RoboDK station: Car_Painting_Model .rdk

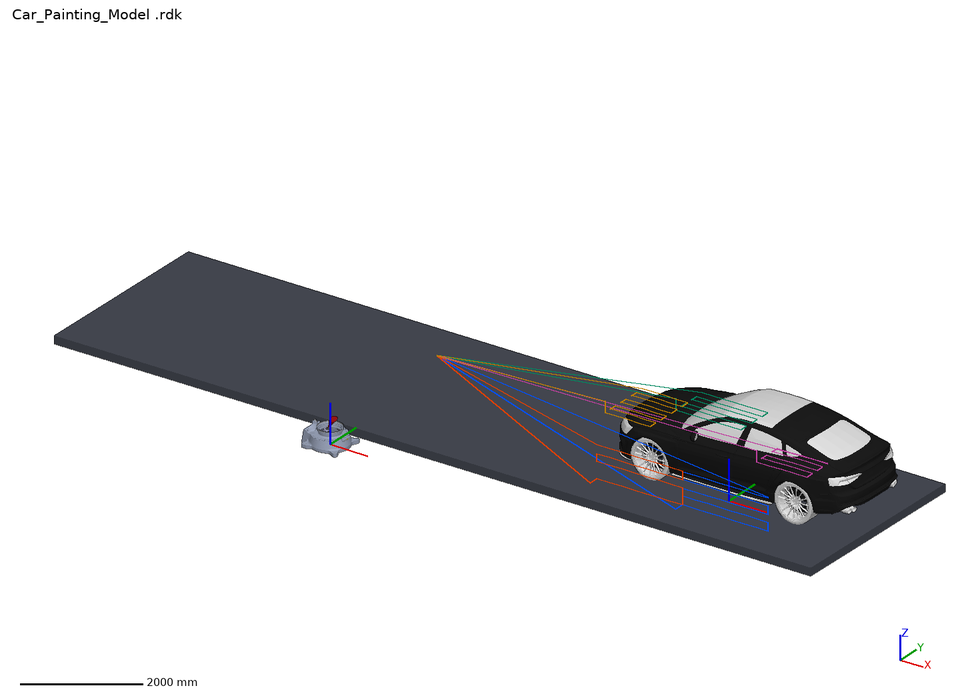
[picture v0: the station drawn from its stored meshes, robots at their saved joint values, targets as dots, program paths as lines]
Station Car_Painting_Model  (saved by RoboDK 6.0.6). Poses are relative to the parent item; angles as X-Y-Z fixed-axis rotations.
Station parameters (name, value as stored): LIN64
  - frame Comau Smart5 NJ 130-2.6 Base at (-637.82, 0, 0) mm
    - robot Comau Smart5 NJ 130-2.6: 6 axes, payload 130 kg, reach 2616 mm, repeatability 0.07 mm, weight 1050 kg
        joint limits [-180, -75, -351, -280, -120, -720] to [180, 95, 170, 280, 120, 720]; home [0, 0, -90, 0, 0, 0]; saved at [0, 0, -90, 0, 0, 0]
      - tool Generic Paint Sprayer, TCP at (50, 0, 450) mm, rotated rx 0 ry 30 rz 0 deg, size 277.6 x 203.2 x 501.7 mm
  - frame CarFrame at (5862.18, 2000, 0) mm
    - object CAN_CAR_BLEND_V12 at (230.98, 0, 65.42) mm, rotated rx 80 ry 0 rz 90 deg, size 2096.9 x 1491.7 x 4800 mm, geometry from CAN_CAR_BLEND_V12.glb
    - target CHK_Nose (Cartesian target) at (2400, 0, 600) mm; joints [0, 0, -90, 0, 0, 0] of Comau Smart5 NJ 130-2.6
    - target CHK_Tail (Cartesian target) at (-2400, 0, 600) mm; joints [0, 0, -90, 0, 0, 0] of Comau Smart5 NJ 130-2.6
    - target CHK_Left_door (Cartesian target) at (0, 1048.43, 800) mm; joints [0, 0, -90, 0, 0, 0] of Comau Smart5 NJ 130-2.6
    - target CHK_Right_door (Cartesian target) at (0, -1048.43, 800) mm; joints [0, 0, -90, 0, 0, 0] of Comau Smart5 NJ 130-2.6
    - target CHK_Roof (Cartesian target) at (0, 0, 1491.68) mm; joints [0, 0, -90, 0, 0, 0] of Comau Smart5 NJ 130-2.6
    - target P_Home (joint target) at (-4384.42, -2000, 2190) mm, rotated rx 180 ry 60 rz 180 deg; joints [0, 0, -90, 0, 0, 0] of Comau Smart5 NJ 130-2.6
    - target P_Right_Front_J_approach (Cartesian target) at (0, -1498.5, 450) mm, rotated rx -90 ry 0 rz 0 deg; joints [0, 0, -90, 0, 0, 0] of Comau Smart5 NJ 130-2.6
    - target P_Right_Front_J_p00_w00 (Cartesian target) at (0, -1298.5, 450) mm, rotated rx -90 ry 0 rz 0 deg; joints [0, 0, -90, 0, 0, 0] of Comau Smart5 NJ 130-2.6
    - target P_Right_Front_J_p00_w01 (Cartesian target) at (242.86, -1298.5, 450) mm, rotated rx -90 ry 0 rz 0 deg; joints [0, 0, -90, 0, 0, 0] of Comau Smart5 NJ 130-2.6
    - target P_Right_Front_J_p00_w02 (Cartesian target) at (485.71, -1298.5, 450) mm, rotated rx -90 ry 0 rz 0 deg; joints [0, 0, -90, 0, 0, 0] of Comau Smart5 NJ 130-2.6
    - target P_Right_Front_J_p00_w03 (Cartesian target) at (728.57, -1298.5, 450) mm, rotated rx -90 ry 0 rz 0 deg; joints [0, 0, -90, 0, 0, 0] of Comau Smart5 NJ 130-2.6
    - target P_Right_Front_J_p00_w04 (Cartesian target) at (971.43, -1298.5, 450) mm, rotated rx -90 ry 0 rz 0 deg; joints [0, 0, -90, 0, 0, 0] of Comau Smart5 NJ 130-2.6
    - target P_Right_Front_J_p00_w05 (Cartesian target) at (1214.29, -1298.5, 450) mm, rotated rx -90 ry 0 rz 0 deg; joints [0, 0, -90, 0, 0, 0] of Comau Smart5 NJ 130-2.6
    - target P_Right_Front_J_p00_w06 (Cartesian target) at (1457.14, -1298.5, 450) mm, rotated rx -90 ry 0 rz 0 deg; joints [0, 0, -90, 0, 0, 0] of Comau Smart5 NJ 130-2.6
    - target P_Right_Front_J_p00_w07 (Cartesian target) at (1700, -1298.5, 450) mm, rotated rx -90 ry 0 rz 0 deg; joints [0, 0, -90, 0, 0, 0] of Comau Smart5 NJ 130-2.6
    - target P_Right_Front_J_p01_w00 (Cartesian target) at (1700, -1298.5, 600) mm, rotated rx 90 ry 0 rz 180 deg; joints [0, 0, -90, 0, 0, 0] of Comau Smart5 NJ 130-2.6
    - target P_Right_Front_J_p01_w01 (Cartesian target) at (1457.14, -1298.5, 600) mm, rotated rx 90 ry 0 rz 180 deg; joints [0, 0, -90, 0, 0, 0] of Comau Smart5 NJ 130-2.6
    - target P_Right_Front_J_p01_w02 (Cartesian target) at (1214.29, -1298.5, 600) mm, rotated rx 90 ry 0 rz 180 deg; joints [0, 0, -90, 0, 0, 0] of Comau Smart5 NJ 130-2.6
    - target P_Right_Front_J_p01_w03 (Cartesian target) at (971.43, -1298.5, 600) mm, rotated rx 90 ry 0 rz 180 deg; joints [0, 0, -90, 0, 0, 0] of Comau Smart5 NJ 130-2.6
    - target P_Right_Front_J_p01_w04 (Cartesian target) at (728.57, -1298.5, 600) mm, rotated rx 90 ry 0 rz 180 deg; joints [0, 0, -90, 0, 0, 0] of Comau Smart5 NJ 130-2.6
    - target P_Right_Front_J_p01_w05 (Cartesian target) at (485.71, -1298.5, 600) mm, rotated rx 90 ry 0 rz 180 deg; joints [0, 0, -90, 0, 0, 0] of Comau Smart5 NJ 130-2.6
    - target P_Right_Front_J_p01_w06 (Cartesian target) at (242.86, -1298.5, 600) mm, rotated rx 90 ry 0 rz 180 deg; joints [0, 0, -90, 0, 0, 0] of Comau Smart5 NJ 130-2.6
    - target P_Right_Front_J_p01_w07 (Cartesian target) at (0, -1298.5, 600) mm, rotated rx 90 ry 0 rz 180 deg; joints [0, 0, -90, 0, 0, 0] of Comau Smart5 NJ 130-2.6
    - target P_Right_Front_J_p02_w00 (Cartesian target) at (0, -1298.5, 750) mm, rotated rx -90 ry 0 rz 0 deg; joints [0, 0, -90, 0, 0, 0] of Comau Smart5 NJ 130-2.6
    - target P_Right_Front_J_p02_w01 (Cartesian target) at (242.86, -1298.5, 750) mm, rotated rx -90 ry 0 rz 0 deg; joints [0, 0, -90, 0, 0, 0] of Comau Smart5 NJ 130-2.6
    - target P_Right_Front_J_p02_w02 (Cartesian target) at (485.71, -1298.5, 750) mm, rotated rx -90 ry 0 rz 0 deg; joints [0, 0, -90, 0, 0, 0] of Comau Smart5 NJ 130-2.6
    - target P_Right_Front_J_p02_w03 (Cartesian target) at (728.57, -1298.5, 750) mm, rotated rx -90 ry 0 rz 0 deg; joints [0, 0, -90, 0, 0, 0] of Comau Smart5 NJ 130-2.6
    - target P_Right_Front_J_p02_w04 (Cartesian target) at (971.43, -1298.5, 750) mm, rotated rx -90 ry 0 rz 0 deg; joints [0, 0, -90, 0, 0, 0] of Comau Smart5 NJ 130-2.6
    - target P_Right_Front_J_p02_w05 (Cartesian target) at (1214.29, -1298.5, 750) mm, rotated rx -90 ry 0 rz 0 deg; joints [0, 0, -90, 0, 0, 0] of Comau Smart5 NJ 130-2.6
    - target P_Right_Front_J_p02_w06 (Cartesian target) at (1457.14, -1298.5, 750) mm, rotated rx -90 ry 0 rz 0 deg; joints [0, 0, -90, 0, 0, 0] of Comau Smart5 NJ 130-2.6
    - target P_Right_Front_J_p02_w07 (Cartesian target) at (1700, -1298.5, 750) mm, rotated rx -90 ry 0 rz 0 deg; joints [0, 0, -90, 0, 0, 0] of Comau Smart5 NJ 130-2.6
    - target P_Right_Front_J_p03_w00 (Cartesian target) at (1700, -1298.5, 900) mm, rotated rx 90 ry 0 rz 180 deg; joints [0, 0, -90, 0, 0, 0] of Comau Smart5 NJ 130-2.6
    - target P_Right_Front_J_p03_w01 (Cartesian target) at (1457.14, -1298.5, 900) mm, rotated rx 90 ry 0 rz 180 deg; joints [0, 0, -90, 0, 0, 0] of Comau Smart5 NJ 130-2.6
    - target P_Right_Front_J_p03_w02 (Cartesian target) at (1214.29, -1298.5, 900) mm, rotated rx 90 ry 0 rz 180 deg; joints [0, 0, -90, 0, 0, 0] of Comau Smart5 NJ 130-2.6
    - target P_Right_Front_J_p03_w03 (Cartesian target) at (971.43, -1298.5, 900) mm, rotated rx 90 ry 0 rz 180 deg; joints [0, 0, -90, 0, 0, 0] of Comau Smart5 NJ 130-2.6
    - target P_Right_Front_J_p03_w04 (Cartesian target) at (728.57, -1298.5, 900) mm, rotated rx 90 ry 0 rz 180 deg; joints [0, 0, -90, 0, 0, 0] of Comau Smart5 NJ 130-2.6
    - target P_Right_Front_J_p03_w05 (Cartesian target) at (485.71, -1298.5, 900) mm, rotated rx 90 ry 0 rz 180 deg; joints [0, 0, -90, 0, 0, 0] of Comau Smart5 NJ 130-2.6
    - target P_Right_Front_J_p03_w06 (Cartesian target) at (242.86, -1298.5, 900) mm, rotated rx 90 ry 0 rz 180 deg; joints [0, 0, -90, 0, 0, 0] of Comau Smart5 NJ 130-2.6
    - target P_Right_Front_J_p03_w07 (Cartesian target) at (0, -1298.5, 900) mm, rotated rx 90 ry 0 rz 180 deg; joints [0, 0, -90, 0, 0, 0] of Comau Smart5 NJ 130-2.6
    - target P_Right_Front_J_p04_w00 (Cartesian target) at (0, -1298.5, 1050) mm, rotated rx -90 ry 0 rz 0 deg; joints [0, 0, -90, 0, 0, 0] of Comau Smart5 NJ 130-2.6
    - target P_Right_Front_J_p04_w01 (Cartesian target) at (242.86, -1298.5, 1050) mm, rotated rx -90 ry 0 rz 0 deg; joints [0, 0, -90, 0, 0, 0] of Comau Smart5 NJ 130-2.6
    - target P_Right_Front_J_p04_w02 (Cartesian target) at (485.71, -1298.5, 1050) mm, rotated rx -90 ry 0 rz 0 deg; joints [0, 0, -90, 0, 0, 0] of Comau Smart5 NJ 130-2.6
    - target P_Right_Front_J_p04_w03 (Cartesian target) at (728.57, -1298.5, 1050) mm, rotated rx -90 ry 0 rz 0 deg; joints [0, 0, -90, 0, 0, 0] of Comau Smart5 NJ 130-2.6
    - target P_Right_Front_J_p04_w04 (Cartesian target) at (971.43, -1298.5, 1050) mm, rotated rx -90 ry 0 rz 0 deg; joints [0, 0, -90, 0, 0, 0] of Comau Smart5 NJ 130-2.6
    - target P_Right_Front_J_p04_w05 (Cartesian target) at (1214.29, -1298.5, 1050) mm, rotated rx -90 ry 0 rz 0 deg; joints [0, 0, -90, 0, 0, 0] of Comau Smart5 NJ 130-2.6
    - target P_Right_Front_J_p04_w06 (Cartesian target) at (1457.14, -1298.5, 1050) mm, rotated rx -90 ry 0 rz 0 deg; joints [0, 0, -90, 0, 0, 0] of Comau Smart5 NJ 130-2.6
    - target P_Right_Front_J_p04_w07 (Cartesian target) at (1700, -1298.5, 1050) mm, rotated rx -90 ry 0 rz 0 deg; joints [0, 0, -90, 0, 0, 0] of Comau Smart5 NJ 130-2.6
    - target P_Right_Rear_J_approach (Cartesian target) at (-1700, -1498.5, 450) mm, rotated rx -90 ry 0 rz 0 deg; joints [-106.937, 43.545, -212.911, 92.647, 99.906, 63.406] of Comau Smart5 NJ 130-2.6
    - target P_Right_Rear_J_p00_w00 (Cartesian target) at (-1700, -1298.5, 450) mm, rotated rx -90 ry 0 rz 0 deg; joints [-106.937, 43.545, -212.911, 92.647, 99.906, 63.406] of Comau Smart5 NJ 130-2.6
    - target P_Right_Rear_J_p00_w01 (Cartesian target) at (-1457.14, -1298.5, 450) mm, rotated rx -90 ry 0 rz 0 deg; joints [-106.937, 43.545, -212.911, 92.647, 99.906, 63.406] of Comau Smart5 NJ 130-2.6
    - target P_Right_Rear_J_p00_w02 (Cartesian target) at (-1214.29, -1298.5, 450) mm, rotated rx -90 ry 0 rz 0 deg; joints [-106.937, 43.545, -212.911, 92.647, 99.906, 63.406] of Comau Smart5 NJ 130-2.6
    - target P_Right_Rear_J_p00_w03 (Cartesian target) at (-971.43, -1298.5, 450) mm, rotated rx -90 ry 0 rz 0 deg; joints [-106.937, 43.545, -212.911, 92.647, 99.906, 63.406] of Comau Smart5 NJ 130-2.6
    - target P_Right_Rear_J_p00_w04 (Cartesian target) at (-728.57, -1298.5, 450) mm, rotated rx -90 ry 0 rz 0 deg; joints [-106.937, 43.545, -212.911, 92.647, 99.906, 63.406] of Comau Smart5 NJ 130-2.6
    - target P_Right_Rear_J_p00_w05 (Cartesian target) at (-485.71, -1298.5, 450) mm, rotated rx -90 ry 0 rz 0 deg; joints [-106.937, 43.545, -212.911, 92.647, 99.906, 63.406] of Comau Smart5 NJ 130-2.6
    - target P_Right_Rear_J_p00_w06 (Cartesian target) at (-242.86, -1298.5, 450) mm, rotated rx -90 ry 0 rz 0 deg; joints [-106.937, 43.545, -212.911, 92.647, 99.906, 63.406] of Comau Smart5 NJ 130-2.6
    - target P_Right_Rear_J_p00_w07 (Cartesian target) at (0, -1298.5, 450) mm, rotated rx -90 ry 0 rz 0 deg; joints [-106.937, 43.545, -212.911, 92.647, 99.906, 63.406] of Comau Smart5 NJ 130-2.6
    - target P_Right_Rear_J_p01_w00 (Cartesian target) at (0, -1298.5, 750) mm, rotated rx -90 ry 0 rz 0 deg; joints [-106.937, 43.545, -212.911, 92.647, 99.906, 63.406] of Comau Smart5 NJ 130-2.6
    - target P_Right_Rear_J_p01_w01 (Cartesian target) at (-242.86, -1298.5, 750) mm, rotated rx -90 ry 0 rz 0 deg; joints [-106.937, 43.545, -212.911, 92.647, 99.906, 63.406] of Comau Smart5 NJ 130-2.6
    - target P_Right_Rear_J_p01_w02 (Cartesian target) at (-485.71, -1298.5, 750) mm, rotated rx -90 ry 0 rz 0 deg; joints [-106.937, 43.545, -212.911, 92.647, 99.906, 63.406] of Comau Smart5 NJ 130-2.6
    - target P_Right_Rear_J_p01_w03 (Cartesian target) at (-728.57, -1298.5, 750) mm, rotated rx -90 ry 0 rz 0 deg; joints [-106.937, 43.545, -212.911, 92.647, 99.906, 63.406] of Comau Smart5 NJ 130-2.6
    - target P_Right_Rear_J_p01_w04 (Cartesian target) at (-971.43, -1298.5, 750) mm, rotated rx -90 ry 0 rz 0 deg; joints [-106.937, 43.545, -212.911, 92.647, 99.906, 63.406] of Comau Smart5 NJ 130-2.6
    - target P_Right_Rear_J_p01_w05 (Cartesian target) at (-1214.29, -1298.5, 750) mm, rotated rx -90 ry 0 rz 0 deg; joints [-106.937, 43.545, -212.911, 92.647, 99.906, 63.406] of Comau Smart5 NJ 130-2.6
    - target P_Right_Rear_J_p01_w06 (Cartesian target) at (-1457.14, -1298.5, 750) mm, rotated rx -90 ry 0 rz 0 deg; joints [-106.937, 43.545, -212.911, 92.647, 99.906, 63.406] of Comau Smart5 NJ 130-2.6
    - target P_Right_Rear_J_p01_w07 (Cartesian target) at (-1700, -1298.5, 750) mm, rotated rx -90 ry 0 rz 0 deg; joints [-106.937, 43.545, -212.911, 92.647, 99.906, 63.406] of Comau Smart5 NJ 130-2.6
    - target P_Right_Rear_J_p02_w00 (Cartesian target) at (-1700, -1298.5, 900) mm, rotated rx 90 ry 0 rz 180 deg; joints [-106.937, 43.545, -212.911, 92.647, 99.906, 63.406] of Comau Smart5 NJ 130-2.6
    - target P_Right_Rear_J_p02_w01 (Cartesian target) at (-1457.14, -1298.5, 900) mm, rotated rx 90 ry 0 rz 180 deg; joints [-106.937, 43.545, -212.911, 92.647, 99.906, 63.406] of Comau Smart5 NJ 130-2.6
    - target P_Right_Rear_J_p02_w02 (Cartesian target) at (-1214.29, -1298.5, 900) mm, rotated rx 90 ry 0 rz 180 deg; joints [-106.937, 43.545, -212.911, 92.647, 99.906, 63.406] of Comau Smart5 NJ 130-2.6
    - target P_Right_Rear_J_p02_w03 (Cartesian target) at (-971.43, -1298.5, 900) mm, rotated rx 90 ry 0 rz 180 deg; joints [-106.937, 43.545, -212.911, 92.647, 99.906, 63.406] of Comau Smart5 NJ 130-2.6
    - target P_Right_Rear_J_p02_w04 (Cartesian target) at (-728.57, -1298.5, 900) mm, rotated rx 90 ry 0 rz 180 deg; joints [-106.937, 43.545, -212.911, 92.647, 99.906, 63.406] of Comau Smart5 NJ 130-2.6
    - target P_Right_Rear_J_p02_w05 (Cartesian target) at (-485.71, -1298.5, 900) mm, rotated rx 90 ry 0 rz 180 deg; joints [-106.937, 43.545, -212.911, 92.647, 99.906, 63.406] of Comau Smart5 NJ 130-2.6
    - target P_Right_Rear_J_p02_w06 (Cartesian target) at (-242.86, -1298.5, 900) mm, rotated rx 90 ry 0 rz 180 deg; joints [-106.937, 43.545, -212.911, 92.647, 99.906, 63.406] of Comau Smart5 NJ 130-2.6
    - target P_Right_Rear_J_p02_w07 (Cartesian target) at (0, -1298.5, 900) mm, rotated rx 90 ry 0 rz 180 deg; joints [-106.937, 43.545, -212.911, 92.647, 99.906, 63.406] of Comau Smart5 NJ 130-2.6
    - target P_Right_Rear_J_p03_w00 (Cartesian target) at (0, -1298.5, 1050) mm, rotated rx -90 ry 0 rz 0 deg; joints [-106.937, 43.545, -212.911, 92.647, 99.906, 63.406] of Comau Smart5 NJ 130-2.6
    - target P_Right_Rear_J_p03_w01 (Cartesian target) at (-242.86, -1298.5, 1050) mm, rotated rx -90 ry 0 rz 0 deg; joints [-106.937, 43.545, -212.911, 92.647, 99.906, 63.406] of Comau Smart5 NJ 130-2.6
    - target P_Right_Rear_J_p03_w02 (Cartesian target) at (-485.71, -1298.5, 1050) mm, rotated rx -90 ry 0 rz 0 deg; joints [-106.937, 43.545, -212.911, 92.647, 99.906, 63.406] of Comau Smart5 NJ 130-2.6
    - target P_Right_Rear_J_p03_w03 (Cartesian target) at (-728.57, -1298.5, 1050) mm, rotated rx -90 ry 0 rz 0 deg; joints [-106.937, 43.545, -212.911, 92.647, 99.906, 63.406] of Comau Smart5 NJ 130-2.6
    - target P_Right_Rear_J_p03_w04 (Cartesian target) at (-971.43, -1298.5, 1050) mm, rotated rx -90 ry 0 rz 0 deg; joints [-106.937, 43.545, -212.911, 92.647, 99.906, 63.406] of Comau Smart5 NJ 130-2.6
    - target P_Right_Rear_J_p03_w05 (Cartesian target) at (-1214.29, -1298.5, 1050) mm, rotated rx -90 ry 0 rz 0 deg; joints [-106.937, 43.545, -212.911, 92.647, 99.906, 63.406] of Comau Smart5 NJ 130-2.6
    - target P_Right_Rear_J_p03_w06 (Cartesian target) at (-1457.14, -1298.5, 1050) mm, rotated rx -90 ry 0 rz 0 deg; joints [-106.937, 43.545, -212.911, 92.647, 99.906, 63.406] of Comau Smart5 NJ 130-2.6
    - target P_Right_Rear_J_p03_w07 (Cartesian target) at (-1700, -1298.5, 1050) mm, rotated rx -90 ry 0 rz 0 deg; joints [-106.937, 43.545, -212.911, 92.647, 99.906, 63.406] of Comau Smart5 NJ 130-2.6
    - target P_Roof_J_approach (Cartesian target) at (-600, -648.5, 1942) mm, rotated rx 180 ry 0 rz 0 deg; joints [0, 0, -90, 0, 0, 0] of Comau Smart5 NJ 130-2.6
    - target P_Roof_J_p00_w00 (Cartesian target) at (-600, -648.5, 1742) mm, rotated rx 180 ry 0 rz 0 deg; joints [0, 0, -90, 0, 0, 0] of Comau Smart5 NJ 130-2.6
    - target P_Roof_J_p00_w01 (Cartesian target) at (-383.33, -648.5, 1742) mm, rotated rx 180 ry 0 rz 0 deg; joints [0, 0, -90, 0, 0, 0] of Comau Smart5 NJ 130-2.6
    - target P_Roof_J_p00_w02 (Cartesian target) at (-166.67, -648.5, 1742) mm, rotated rx 180 ry 0 rz 0 deg; joints [0, 0, -90, 0, 0, 0] of Comau Smart5 NJ 130-2.6
    - target P_Roof_J_p00_w03 (Cartesian target) at (50, -648.5, 1742) mm, rotated rx 180 ry 0 rz 0 deg; joints [0, 0, -90, 0, 0, 0] of Comau Smart5 NJ 130-2.6
    - target P_Roof_J_p00_w04 (Cartesian target) at (266.67, -648.5, 1742) mm, rotated rx 180 ry 0 rz 0 deg; joints [0, 0, -90, 0, 0, 0] of Comau Smart5 NJ 130-2.6
    - target P_Roof_J_p00_w05 (Cartesian target) at (483.33, -648.5, 1742) mm, rotated rx 180 ry 0 rz 0 deg; joints [0, 0, -90, 0, 0, 0] of Comau Smart5 NJ 130-2.6
    - target P_Roof_J_p00_w06 (Cartesian target) at (700, -648.5, 1742) mm, rotated rx 180 ry 0 rz 0 deg; joints [0, 0, -90, 0, 0, 0] of Comau Smart5 NJ 130-2.6
    - target P_Roof_J_p01_w00 (Cartesian target) at (700, -498.5, 1742) mm, rotated rx 180 ry 0 rz 180 deg; joints [0, 0, -90, 0, 0, 0] of Comau Smart5 NJ 130-2.6
    - target P_Roof_J_p01_w01 (Cartesian target) at (483.33, -498.5, 1742) mm, rotated rx 180 ry 0 rz 180 deg; joints [0, 0, -90, 0, 0, 0] of Comau Smart5 NJ 130-2.6
    - target P_Roof_J_p01_w02 (Cartesian target) at (266.67, -498.5, 1742) mm, rotated rx 180 ry 0 rz 180 deg; joints [0, 0, -90, 0, 0, 0] of Comau Smart5 NJ 130-2.6
    - target P_Roof_J_p01_w03 (Cartesian target) at (50, -498.5, 1742) mm, rotated rx 180 ry 0 rz 180 deg; joints [0, 0, -90, 0, 0, 0] of Comau Smart5 NJ 130-2.6
    - target P_Roof_J_p01_w04 (Cartesian target) at (-166.67, -498.5, 1742) mm, rotated rx 180 ry 0 rz 180 deg; joints [0, 0, -90, 0, 0, 0] of Comau Smart5 NJ 130-2.6
    - target P_Roof_J_p01_w05 (Cartesian target) at (-383.33, -498.5, 1742) mm, rotated rx 180 ry 0 rz 180 deg; joints [0, 0, -90, 0, 0, 0] of Comau Smart5 NJ 130-2.6
    - target P_Roof_J_p01_w06 (Cartesian target) at (-600, -498.5, 1742) mm, rotated rx 180 ry 0 rz 180 deg; joints [0, 0, -90, 0, 0, 0] of Comau Smart5 NJ 130-2.6
    - target P_Roof_J_p02_w00 (Cartesian target) at (-600, -348.5, 1742) mm, rotated rx 180 ry 0 rz 0 deg; joints [0, 0, -90, 0, 0, 0] of Comau Smart5 NJ 130-2.6
    - target P_Roof_J_p02_w01 (Cartesian target) at (-383.33, -348.5, 1742) mm, rotated rx 180 ry 0 rz 0 deg; joints [0, 0, -90, 0, 0, 0] of Comau Smart5 NJ 130-2.6
    - target P_Roof_J_p02_w02 (Cartesian target) at (-166.67, -348.5, 1742) mm, rotated rx 180 ry 0 rz 0 deg; joints [0, 0, -90, 0, 0, 0] of Comau Smart5 NJ 130-2.6
    - target P_Roof_J_p02_w03 (Cartesian target) at (50, -348.5, 1742) mm, rotated rx 180 ry 0 rz 0 deg; joints [0, 0, -90, 0, 0, 0] of Comau Smart5 NJ 130-2.6
    - target P_Roof_J_p02_w04 (Cartesian target) at (266.67, -348.5, 1742) mm, rotated rx 180 ry 0 rz 0 deg; joints [0, 0, -90, 0, 0, 0] of Comau Smart5 NJ 130-2.6
    - target P_Roof_J_p02_w05 (Cartesian target) at (483.33, -348.5, 1742) mm, rotated rx 180 ry 0 rz 0 deg; joints [0, 0, -90, 0, 0, 0] of Comau Smart5 NJ 130-2.6
    - target P_Roof_J_p02_w06 (Cartesian target) at (700, -348.5, 1742) mm, rotated rx 180 ry 0 rz 0 deg; joints [0, 0, -90, 0, 0, 0] of Comau Smart5 NJ 130-2.6
    - target P_Roof_J_p03_w00 (Cartesian target) at (700, -198.5, 1742) mm, rotated rx 180 ry 0 rz 180 deg; joints [0, 0, -90, 0, 0, 0] of Comau Smart5 NJ 130-2.6
    - target P_Roof_J_p03_w01 (Cartesian target) at (483.33, -198.5, 1742) mm, rotated rx 180 ry 0 rz 180 deg; joints [0, 0, -90, 0, 0, 0] of Comau Smart5 NJ 130-2.6
    - target P_Roof_J_p03_w02 (Cartesian target) at (266.67, -198.5, 1742) mm, rotated rx 180 ry 0 rz 180 deg; joints [0, 0, -90, 0, 0, 0] of Comau Smart5 NJ 130-2.6
    - target P_Roof_J_p03_w03 (Cartesian target) at (50, -198.5, 1742) mm, rotated rx 180 ry 0 rz 180 deg; joints [0, 0, -90, 0, 0, 0] of Comau Smart5 NJ 130-2.6
    - target P_Roof_J_p03_w04 (Cartesian target) at (-166.67, -198.5, 1742) mm, rotated rx 180 ry 0 rz 180 deg; joints [0, 0, -90, 0, 0, 0] of Comau Smart5 NJ 130-2.6
    - target P_Roof_J_p03_w05 (Cartesian target) at (-383.33, -198.5, 1742) mm, rotated rx 180 ry 0 rz 180 deg; joints [0, 0, -90, 0, 0, 0] of Comau Smart5 NJ 130-2.6
    - target P_Roof_J_p03_w06 (Cartesian target) at (-600, -198.5, 1742) mm, rotated rx 180 ry 0 rz 180 deg; joints [0, 0, -90, 0, 0, 0] of Comau Smart5 NJ 130-2.6
    - target P_Roof_J_p04_w00 (Cartesian target) at (-600, -48.5, 1742) mm, rotated rx -160 ry 0 rz 0 deg; joints [0, 0, -90, 0, 0, 0] of Comau Smart5 NJ 130-2.6
    - target P_Roof_J_p04_w01 (Cartesian target) at (-383.33, -48.5, 1742) mm, rotated rx -160 ry 0 rz 0 deg; joints [0, 0, -90, 0, 0, 0] of Comau Smart5 NJ 130-2.6
    - target P_Roof_J_p04_w02 (Cartesian target) at (-166.67, -48.5, 1742) mm, rotated rx -160 ry 0 rz 0 deg; joints [0, 0, -90, 0, 0, 0] of Comau Smart5 NJ 130-2.6
    - target P_Roof_J_p04_w03 (Cartesian target) at (50, -48.5, 1742) mm, rotated rx -160 ry 0 rz 0 deg; joints [0, 0, -90, 0, 0, 0] of Comau Smart5 NJ 130-2.6
    - target P_Roof_J_p04_w04 (Cartesian target) at (266.67, -48.5, 1742) mm, rotated rx -160 ry 0 rz 0 deg; joints [0, 0, -90, 0, 0, 0] of Comau Smart5 NJ 130-2.6
    - target P_Roof_J_p04_w05 (Cartesian target) at (483.33, -48.5, 1742) mm, rotated rx -160 ry 0 rz 0 deg; joints [0, 0, -90, 0, 0, 0] of Comau Smart5 NJ 130-2.6
    - target P_Roof_J_p04_w06 (Cartesian target) at (700, -48.5, 1742) mm, rotated rx -160 ry 0 rz 0 deg; joints [0, 0, -90, 0, 0, 0] of Comau Smart5 NJ 130-2.6
    - target P_Roof_J_p05_w00 (Cartesian target) at (700, 101.5, 1742) mm, rotated rx 160 ry 0 rz 180 deg; joints [0, 0, -90, 0, 0, 0] of Comau Smart5 NJ 130-2.6
    - target P_Roof_J_p05_w01 (Cartesian target) at (483.33, 101.5, 1742) mm, rotated rx 160 ry 0 rz 180 deg; joints [0, 0, -90, 0, 0, 0] of Comau Smart5 NJ 130-2.6
    - target P_Roof_J_p05_w02 (Cartesian target) at (266.67, 101.5, 1742) mm, rotated rx 160 ry 0 rz 180 deg; joints [0, 0, -90, 0, 0, 0] of Comau Smart5 NJ 130-2.6
    - target P_Roof_J_p05_w03 (Cartesian target) at (50, 101.5, 1742) mm, rotated rx 160 ry 0 rz 180 deg; joints [0, 0, -90, 0, 0, 0] of Comau Smart5 NJ 130-2.6
    - target P_Roof_J_p05_w04 (Cartesian target) at (-166.67, 101.5, 1742) mm, rotated rx 160 ry 0 rz 180 deg; joints [0, 0, -90, 0, 0, 0] of Comau Smart5 NJ 130-2.6
    - target P_Roof_J_p05_w05 (Cartesian target) at (-383.33, 101.5, 1742) mm, rotated rx 160 ry 0 rz 180 deg; joints [0, 0, -90, 0, 0, 0] of Comau Smart5 NJ 130-2.6
    - target P_Roof_J_p05_w06 (Cartesian target) at (-600, 101.5, 1742) mm, rotated rx 160 ry 0 rz 180 deg; joints [0, 0, -90, 0, 0, 0] of Comau Smart5 NJ 130-2.6
    - target P_Hood_J_approach (Cartesian target) at (1000, -648.5, 1450) mm, rotated rx 180 ry 0 rz -180 deg; joints [-82.567, 85.196, -51.536, -34.414, 109.08, 85.646] of Comau Smart5 NJ 130-2.6
    - target P_Hood_J_p00_w00 (Cartesian target) at (1000, -648.5, 1250) mm, rotated rx 180 ry 0 rz -180 deg; joints [-82.567, 85.196, -51.536, -34.414, 109.08, 85.646] of Comau Smart5 NJ 130-2.6
    - target P_Hood_J_p00_w01 (Cartesian target) at (1250, -648.5, 1250) mm, rotated rx 180 ry 0 rz -180 deg; joints [-82.567, 85.196, -51.536, -34.414, 109.08, 85.646] of Comau Smart5 NJ 130-2.6
    - target P_Hood_J_p00_w02 (Cartesian target) at (1500, -648.5, 1250) mm, rotated rx 180 ry 0 rz -180 deg; joints [-82.567, 85.196, -51.536, -34.414, 109.08, 85.646] of Comau Smart5 NJ 130-2.6
    - target P_Hood_J_p00_w03 (Cartesian target) at (1750, -648.5, 1250) mm, rotated rx 180 ry 0 rz -180 deg; joints [-82.567, 85.196, -51.536, -34.414, 109.08, 85.646] of Comau Smart5 NJ 130-2.6
    - target P_Hood_J_p00_w04 (Cartesian target) at (2000, -648.5, 1250) mm, rotated rx 180 ry 0 rz -180 deg; joints [-82.567, 85.196, -51.536, -34.414, 109.08, 85.646] of Comau Smart5 NJ 130-2.6
    - target P_Hood_J_p01_w00 (Cartesian target) at (2000, -498.5, 1250) mm, rotated rx 180 ry 0 rz 0 deg; joints [-82.567, 85.196, -51.536, -34.414, 109.08, 85.646] of Comau Smart5 NJ 130-2.6
    - target P_Hood_J_p01_w01 (Cartesian target) at (1750, -498.5, 1250) mm, rotated rx 180 ry 0 rz 0 deg; joints [-82.567, 85.196, -51.536, -34.414, 109.08, 85.646] of Comau Smart5 NJ 130-2.6
    - target P_Hood_J_p01_w02 (Cartesian target) at (1500, -498.5, 1250) mm, rotated rx 180 ry 0 rz 0 deg; joints [-82.567, 85.196, -51.536, -34.414, 109.08, 85.646] of Comau Smart5 NJ 130-2.6
    - target P_Hood_J_p01_w03 (Cartesian target) at (1250, -498.5, 1250) mm, rotated rx 180 ry 0 rz 0 deg; joints [-82.567, 85.196, -51.536, -34.414, 109.08, 85.646] of Comau Smart5 NJ 130-2.6
    - target P_Hood_J_p01_w04 (Cartesian target) at (1000, -498.5, 1250) mm, rotated rx 180 ry 0 rz 0 deg; joints [-82.567, 85.196, -51.536, -34.414, 109.08, 85.646] of Comau Smart5 NJ 130-2.6
    - target P_Hood_J_p02_w00 (Cartesian target) at (1000, -348.5, 1250) mm, rotated rx 180 ry 0 rz -180 deg; joints [-82.567, 85.196, -51.536, -34.414, 109.08, 85.646] of Comau Smart5 NJ 130-2.6
    - target P_Hood_J_p02_w01 (Cartesian target) at (1250, -348.5, 1250) mm, rotated rx 180 ry 0 rz -180 deg; joints [-82.567, 85.196, -51.536, -34.414, 109.08, 85.646] of Comau Smart5 NJ 130-2.6
    - target P_Hood_J_p02_w02 (Cartesian target) at (1500, -348.5, 1250) mm, rotated rx 180 ry 0 rz -180 deg; joints [-82.567, 85.196, -51.536, -34.414, 109.08, 85.646] of Comau Smart5 NJ 130-2.6
    - target P_Hood_J_p02_w03 (Cartesian target) at (1750, -348.5, 1250) mm, rotated rx 180 ry 0 rz -180 deg; joints [-82.567, 85.196, -51.536, -34.414, 109.08, 85.646] of Comau Smart5 NJ 130-2.6
    - target P_Hood_J_p02_w04 (Cartesian target) at (2000, -348.5, 1250) mm, rotated rx 180 ry 0 rz -180 deg; joints [-82.567, 85.196, -51.536, -34.414, 109.08, 85.646] of Comau Smart5 NJ 130-2.6
    - target P_Hood_J_p03_w00 (Cartesian target) at (2000, -198.5, 1250) mm, rotated rx 180 ry 0 rz 0 deg; joints [-82.567, 85.196, -51.536, -34.414, 109.08, 85.646] of Comau Smart5 NJ 130-2.6
    - target P_Hood_J_p03_w01 (Cartesian target) at (1750, -198.5, 1250) mm, rotated rx 180 ry 0 rz 0 deg; joints [-82.567, 85.196, -51.536, -34.414, 109.08, 85.646] of Comau Smart5 NJ 130-2.6
    - target P_Hood_J_p03_w02 (Cartesian target) at (1500, -198.5, 1250) mm, rotated rx 180 ry 0 rz 0 deg; joints [-82.567, 85.196, -51.536, -34.414, 109.08, 85.646] of Comau Smart5 NJ 130-2.6
    - target P_Hood_J_p03_w03 (Cartesian target) at (1250, -198.5, 1250) mm, rotated rx 180 ry 0 rz 0 deg; joints [-82.567, 85.196, -51.536, -34.414, 109.08, 85.646] of Comau Smart5 NJ 130-2.6
    - target P_Hood_J_p03_w04 (Cartesian target) at (1000, -198.5, 1250) mm, rotated rx 180 ry 0 rz 0 deg; joints [-82.567, 85.196, -51.536, -34.414, 109.08, 85.646] of Comau Smart5 NJ 130-2.6
    - target P_Hood_J_p04_w00 (Cartesian target) at (1000, -48.5, 1250) mm, rotated rx 180 ry 0 rz -180 deg; joints [-82.567, 85.196, -51.536, -34.414, 109.08, 85.646] of Comau Smart5 NJ 130-2.6
    - target P_Hood_J_p04_w01 (Cartesian target) at (1250, -48.5, 1250) mm, rotated rx 180 ry 0 rz -180 deg; joints [-82.567, 85.196, -51.536, -34.414, 109.08, 85.646] of Comau Smart5 NJ 130-2.6
    - target P_Hood_J_p04_w02 (Cartesian target) at (1500, -48.5, 1250) mm, rotated rx 180 ry 0 rz -180 deg; joints [-82.567, 85.196, -51.536, -34.414, 109.08, 85.646] of Comau Smart5 NJ 130-2.6
    - target P_Hood_J_p04_w03 (Cartesian target) at (1750, -48.5, 1250) mm, rotated rx 180 ry 0 rz -180 deg; joints [-82.567, 85.196, -51.536, -34.414, 109.08, 85.646] of Comau Smart5 NJ 130-2.6
    - target P_Hood_J_p04_w04 (Cartesian target) at (2000, -48.5, 1250) mm, rotated rx 180 ry 0 rz -180 deg; joints [-82.567, 85.196, -51.536, -34.414, 109.08, 85.646] of Comau Smart5 NJ 130-2.6
    - target P_Trunk_J_approach (Cartesian target) at (-2000, -648.5, 1500) mm, rotated rx 180 ry 0 rz 0 deg; joints [0, 0, -90, 0, 0, 0] of Comau Smart5 NJ 130-2.6
    - target P_Trunk_J_p00_w00 (Cartesian target) at (-2000, -648.5, 1300) mm, rotated rx 180 ry 0 rz 0 deg; joints [0, 0, -90, 0, 0, 0] of Comau Smart5 NJ 130-2.6
    - target P_Trunk_J_p00_w01 (Cartesian target) at (-1775, -648.5, 1300) mm, rotated rx 180 ry 0 rz 0 deg; joints [0, 0, -90, 0, 0, 0] of Comau Smart5 NJ 130-2.6
    - target P_Trunk_J_p00_w02 (Cartesian target) at (-1550, -648.5, 1300) mm, rotated rx 180 ry 0 rz 0 deg; joints [0, 0, -90, 0, 0, 0] of Comau Smart5 NJ 130-2.6
    - target P_Trunk_J_p00_w03 (Cartesian target) at (-1325, -648.5, 1300) mm, rotated rx 180 ry 0 rz 0 deg; joints [0, 0, -90, 0, 0, 0] of Comau Smart5 NJ 130-2.6
    - target P_Trunk_J_p00_w04 (Cartesian target) at (-1100, -648.5, 1300) mm, rotated rx 180 ry 0 rz 0 deg; joints [0, 0, -90, 0, 0, 0] of Comau Smart5 NJ 130-2.6
    - target P_Trunk_J_p01_w00 (Cartesian target) at (-1100, -498.5, 1300) mm, rotated rx 180 ry 0 rz 180 deg; joints [0, 0, -90, 0, 0, 0] of Comau Smart5 NJ 130-2.6
    - target P_Trunk_J_p01_w01 (Cartesian target) at (-1325, -498.5, 1300) mm, rotated rx 180 ry 0 rz 180 deg; joints [0, 0, -90, 0, 0, 0] of Comau Smart5 NJ 130-2.6
    - target P_Trunk_J_p01_w02 (Cartesian target) at (-1550, -498.5, 1300) mm, rotated rx 180 ry 0 rz 180 deg; joints [0, 0, -90, 0, 0, 0] of Comau Smart5 NJ 130-2.6
    - target P_Trunk_J_p01_w03 (Cartesian target) at (-1775, -498.5, 1300) mm, rotated rx 180 ry 0 rz 180 deg; joints [0, 0, -90, 0, 0, 0] of Comau Smart5 NJ 130-2.6
    - target P_Trunk_J_p01_w04 (Cartesian target) at (-2000, -498.5, 1300) mm, rotated rx 180 ry 0 rz 180 deg; joints [0, 0, -90, 0, 0, 0] of Comau Smart5 NJ 130-2.6
    - target P_Trunk_J_p02_w00 (Cartesian target) at (-2000, -348.5, 1300) mm, rotated rx 180 ry 0 rz 0 deg; joints [0, 0, -90, 0, 0, 0] of Comau Smart5 NJ 130-2.6
    - target P_Trunk_J_p02_w01 (Cartesian target) at (-1775, -348.5, 1300) mm, rotated rx 180 ry 0 rz 0 deg; joints [0, 0, -90, 0, 0, 0] of Comau Smart5 NJ 130-2.6
    - target P_Trunk_J_p02_w02 (Cartesian target) at (-1550, -348.5, 1300) mm, rotated rx 180 ry 0 rz 0 deg; joints [0, 0, -90, 0, 0, 0] of Comau Smart5 NJ 130-2.6
    - target P_Trunk_J_p02_w03 (Cartesian target) at (-1325, -348.5, 1300) mm, rotated rx 180 ry 0 rz 0 deg; joints [0, 0, -90, 0, 0, 0] of Comau Smart5 NJ 130-2.6
    - target P_Trunk_J_p02_w04 (Cartesian target) at (-1100, -348.5, 1300) mm, rotated rx 180 ry 0 rz 0 deg; joints [0, 0, -90, 0, 0, 0] of Comau Smart5 NJ 130-2.6
    - target P_Trunk_J_p03_w00 (Cartesian target) at (-1100, -198.5, 1300) mm, rotated rx 180 ry 0 rz 180 deg; joints [0, 0, -90, 0, 0, 0] of Comau Smart5 NJ 130-2.6
    - target P_Trunk_J_p03_w01 (Cartesian target) at (-1325, -198.5, 1300) mm, rotated rx 180 ry 0 rz 180 deg; joints [0, 0, -90, 0, 0, 0] of Comau Smart5 NJ 130-2.6
    - target P_Trunk_J_p03_w02 (Cartesian target) at (-1550, -198.5, 1300) mm, rotated rx 180 ry 0 rz 180 deg; joints [0, 0, -90, 0, 0, 0] of Comau Smart5 NJ 130-2.6
    - target P_Trunk_J_p03_w03 (Cartesian target) at (-1775, -198.5, 1300) mm, rotated rx 180 ry 0 rz 180 deg; joints [0, 0, -90, 0, 0, 0] of Comau Smart5 NJ 130-2.6
    - target P_Trunk_J_p03_w04 (Cartesian target) at (-2000, -198.5, 1300) mm, rotated rx 180 ry 0 rz 180 deg; joints [0, 0, -90, 0, 0, 0] of Comau Smart5 NJ 130-2.6
    - target P_Trunk_J_p04_w00 (Cartesian target) at (-2000, -48.5, 1300) mm, rotated rx 180 ry 0 rz 0 deg; joints [0, 0, -90, 0, 0, 0] of Comau Smart5 NJ 130-2.6
    - target P_Trunk_J_p04_w01 (Cartesian target) at (-1775, -48.5, 1300) mm, rotated rx 180 ry 0 rz 0 deg; joints [0, 0, -90, 0, 0, 0] of Comau Smart5 NJ 130-2.6
    - target P_Trunk_J_p04_w02 (Cartesian target) at (-1550, -48.5, 1300) mm, rotated rx 180 ry 0 rz 0 deg; joints [0, 0, -90, 0, 0, 0] of Comau Smart5 NJ 130-2.6
    - target P_Trunk_J_p04_w03 (Cartesian target) at (-1325, -48.5, 1300) mm, rotated rx 180 ry 0 rz 0 deg; joints [0, 0, -90, 0, 0, 0] of Comau Smart5 NJ 130-2.6
    - target P_Trunk_J_p04_w04 (Cartesian target) at (-1100, -48.5, 1300) mm, rotated rx 180 ry 0 rz 0 deg; joints [0, 0, -90, 0, 0, 0] of Comau Smart5 NJ 130-2.6
    - target P_Trunk_J_p05_w00 (Cartesian target) at (-1100, 101.5, 1300) mm, rotated rx 180 ry 0 rz 180 deg; joints [0, 0, -90, 0, 0, 0] of Comau Smart5 NJ 130-2.6
    - target P_Trunk_J_p05_w01 (Cartesian target) at (-1325, 101.5, 1300) mm, rotated rx 180 ry 0 rz 180 deg; joints [0, 0, -90, 0, 0, 0] of Comau Smart5 NJ 130-2.6
    - target P_Trunk_J_p05_w02 (Cartesian target) at (-1550, 101.5, 1300) mm, rotated rx 180 ry 0 rz 180 deg; joints [0, 0, -90, 0, 0, 0] of Comau Smart5 NJ 130-2.6
    - target P_Trunk_J_p05_w03 (Cartesian target) at (-1775, 101.5, 1300) mm, rotated rx 180 ry 0 rz 180 deg; joints [0, 0, -90, 0, 0, 0] of Comau Smart5 NJ 130-2.6
    - target P_Trunk_J_p05_w04 (Cartesian target) at (-2000, 101.5, 1300) mm, rotated rx 180 ry 0 rz 180 deg; joints [0, 0, -90, 0, 0, 0] of Comau Smart5 NJ 130-2.6
    - target P_Trunk_J_p06_w00 (Cartesian target) at (-2000, 251.5, 1300) mm, rotated rx 180 ry 0 rz 0 deg; joints [0, 0, -90, 0, 0, 0] of Comau Smart5 NJ 130-2.6
    - target P_Trunk_J_p06_w01 (Cartesian target) at (-1775, 251.5, 1300) mm, rotated rx 180 ry 0 rz 0 deg; joints [0, 0, -90, 0, 0, 0] of Comau Smart5 NJ 130-2.6
    - target P_Trunk_J_p06_w02 (Cartesian target) at (-1550, 251.5, 1300) mm, rotated rx 180 ry 0 rz 0 deg; joints [0, 0, -90, 0, 0, 0] of Comau Smart5 NJ 130-2.6
    - target P_Trunk_J_p06_w03 (Cartesian target) at (-1325, 251.5, 1300) mm, rotated rx 180 ry 0 rz 0 deg; joints [0, 0, -90, 0, 0, 0] of Comau Smart5 NJ 130-2.6
    - target P_Trunk_J_p06_w04 (Cartesian target) at (-1100, 251.5, 1300) mm, rotated rx 180 ry 0 rz 0 deg; joints [0, 0, -90, 0, 0, 0] of Comau Smart5 NJ 130-2.6
    - target P_Trunk_J_p07_w00 (Cartesian target) at (-1100, 401.5, 1300) mm, rotated rx 160 ry 0 rz 180 deg; joints [0, 0, -90, 0, 0, 0] of Comau Smart5 NJ 130-2.6
    - target P_Trunk_J_p07_w01 (Cartesian target) at (-1325, 401.5, 1300) mm, rotated rx 160 ry 0 rz 180 deg; joints [0, 0, -90, 0, 0, 0] of Comau Smart5 NJ 130-2.6
    - target P_Trunk_J_p07_w02 (Cartesian target) at (-1550, 401.5, 1300) mm, rotated rx 160 ry 0 rz 180 deg; joints [0, 0, -90, 0, 0, 0] of Comau Smart5 NJ 130-2.6
    - target P_Trunk_J_p07_w03 (Cartesian target) at (-1775, 401.5, 1300) mm, rotated rx 160 ry 0 rz 180 deg; joints [0, 0, -90, 0, 0, 0] of Comau Smart5 NJ 130-2.6
    - target P_Trunk_J_p07_w04 (Cartesian target) at (-2000, 401.5, 1300) mm, rotated rx 160 ry 0 rz 180 deg; joints [0, 0, -90, 0, 0, 0] of Comau Smart5 NJ 130-2.6
  - object Conveyor at (862.18, 2650, -10) mm, size 15000 x 3800 x 150 mm, geometry from conveyor.stl
  - program Paint_Right_Front (45 instructions, listed below)
  - program Paint_Right_Rear (37 instructions, listed below)
  - program Paint_Roof (47 instructions, listed below)
  - program Paint_Hood (30 instructions, listed below)
  - program Paint_Trunk (45 instructions, listed below)
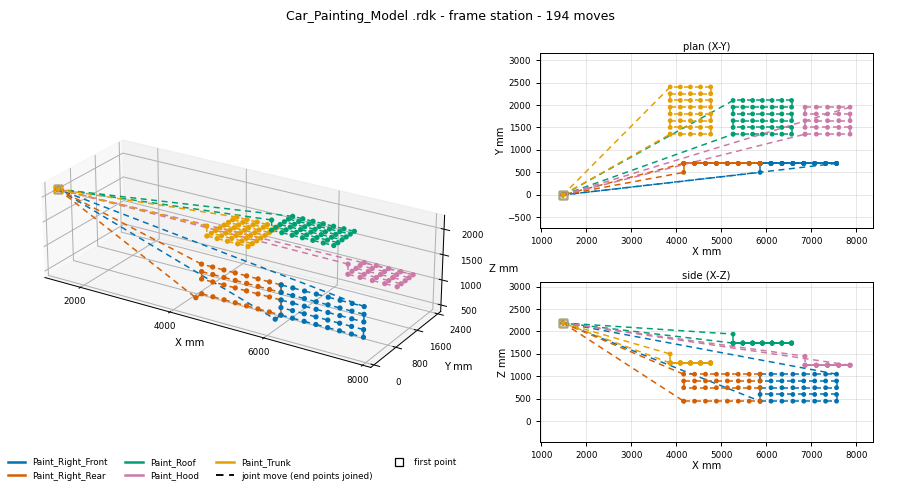
[picture p0: tool path of Car_Painting_Model .rdk in frame station, 194 of 194 moves have a stored position in this frame; points joined in program order, loops and branches not executed]

--- program Paint_Right_Front (robot Comau Smart5 NJ 130-2.6) ---
  Set Ref.: CarFrame
  Set Tool: Generic Paint Sprayer
  MoveJ (P_Home)
  MoveJ (P_Right_Front_J_approach)
  MoveJ (P_Right_Front_J_p00_w00)
  MoveJ (P_Right_Front_J_p00_w01)
  MoveJ (P_Right_Front_J_p00_w02)
  MoveJ (P_Right_Front_J_p00_w03)
  MoveJ (P_Right_Front_J_p00_w04)
  MoveJ (P_Right_Front_J_p00_w05)
  MoveJ (P_Right_Front_J_p00_w06)
  MoveJ (P_Right_Front_J_p00_w07)
  MoveJ (P_Right_Front_J_p01_w00)
  MoveJ (P_Right_Front_J_p01_w01)
  MoveJ (P_Right_Front_J_p01_w02)
  MoveJ (P_Right_Front_J_p01_w03)
  MoveJ (P_Right_Front_J_p01_w04)
  MoveJ (P_Right_Front_J_p01_w05)
  MoveJ (P_Right_Front_J_p01_w06)
  MoveJ (P_Right_Front_J_p01_w07)
  MoveJ (P_Right_Front_J_p02_w00)
  MoveJ (P_Right_Front_J_p02_w01)
  MoveJ (P_Right_Front_J_p02_w02)
  MoveJ (P_Right_Front_J_p02_w03)
  MoveJ (P_Right_Front_J_p02_w04)
  MoveJ (P_Right_Front_J_p02_w05)
  MoveJ (P_Right_Front_J_p02_w06)
  MoveJ (P_Right_Front_J_p02_w07)
  MoveJ (P_Right_Front_J_p03_w00)
  MoveJ (P_Right_Front_J_p03_w01)
  MoveJ (P_Right_Front_J_p03_w02)
  MoveJ (P_Right_Front_J_p03_w03)
  MoveJ (P_Right_Front_J_p03_w04)
  MoveJ (P_Right_Front_J_p03_w05)
  MoveJ (P_Right_Front_J_p03_w06)
  MoveJ (P_Right_Front_J_p03_w07)
  MoveJ (P_Right_Front_J_p04_w00)
  MoveJ (P_Right_Front_J_p04_w01)
  MoveJ (P_Right_Front_J_p04_w02)
  MoveJ (P_Right_Front_J_p04_w03)
  MoveJ (P_Right_Front_J_p04_w04)
  MoveJ (P_Right_Front_J_p04_w05)
  MoveJ (P_Right_Front_J_p04_w06)
  MoveJ (P_Right_Front_J_p04_w07)
  MoveJ (P_Home)

--- program Paint_Right_Rear (robot Comau Smart5 NJ 130-2.6) ---
  Set Ref.: CarFrame
  Set Tool: Generic Paint Sprayer
  MoveJ (P_Home)
  MoveJ (P_Right_Rear_J_approach)
  MoveJ (P_Right_Rear_J_p00_w00)
  MoveJ (P_Right_Rear_J_p00_w01)
  MoveJ (P_Right_Rear_J_p00_w02)
  MoveJ (P_Right_Rear_J_p00_w03)
  MoveJ (P_Right_Rear_J_p00_w04)
  MoveJ (P_Right_Rear_J_p00_w05)
  MoveJ (P_Right_Rear_J_p00_w06)
  MoveJ (P_Right_Rear_J_p00_w07)
  MoveJ (P_Right_Rear_J_p01_w00)
  MoveJ (P_Right_Rear_J_p01_w01)
  MoveJ (P_Right_Rear_J_p01_w02)
  MoveJ (P_Right_Rear_J_p01_w03)
  MoveJ (P_Right_Rear_J_p01_w04)
  MoveJ (P_Right_Rear_J_p01_w05)
  MoveJ (P_Right_Rear_J_p01_w06)
  MoveJ (P_Right_Rear_J_p01_w07)
  MoveJ (P_Right_Rear_J_p02_w00)
  MoveJ (P_Right_Rear_J_p02_w01)
  MoveJ (P_Right_Rear_J_p02_w02)
  MoveJ (P_Right_Rear_J_p02_w03)
  MoveJ (P_Right_Rear_J_p02_w04)
  MoveJ (P_Right_Rear_J_p02_w05)
  MoveJ (P_Right_Rear_J_p02_w06)
  MoveJ (P_Right_Rear_J_p02_w07)
  MoveJ (P_Right_Rear_J_p03_w00)
  MoveJ (P_Right_Rear_J_p03_w01)
  MoveJ (P_Right_Rear_J_p03_w02)
  MoveJ (P_Right_Rear_J_p03_w03)
  MoveJ (P_Right_Rear_J_p03_w04)
  MoveJ (P_Right_Rear_J_p03_w05)
  MoveJ (P_Right_Rear_J_p03_w06)
  MoveJ (P_Right_Rear_J_p03_w07)
  MoveJ (P_Home)

--- program Paint_Roof (robot Comau Smart5 NJ 130-2.6) ---
  Set Ref.: CarFrame
  Set Tool: Generic Paint Sprayer
  MoveJ (P_Home)
  MoveJ (P_Roof_J_approach)
  MoveJ (P_Roof_J_p00_w00)
  MoveJ (P_Roof_J_p00_w01)
  MoveJ (P_Roof_J_p00_w02)
  MoveJ (P_Roof_J_p00_w03)
  MoveJ (P_Roof_J_p00_w04)
  MoveJ (P_Roof_J_p00_w05)
  MoveJ (P_Roof_J_p00_w06)
  MoveJ (P_Roof_J_p01_w00)
  MoveJ (P_Roof_J_p01_w01)
  MoveJ (P_Roof_J_p01_w02)
  MoveJ (P_Roof_J_p01_w03)
  MoveJ (P_Roof_J_p01_w04)
  MoveJ (P_Roof_J_p01_w05)
  MoveJ (P_Roof_J_p01_w06)
  MoveJ (P_Roof_J_p02_w00)
  MoveJ (P_Roof_J_p02_w01)
  MoveJ (P_Roof_J_p02_w02)
  MoveJ (P_Roof_J_p02_w03)
  MoveJ (P_Roof_J_p02_w04)
  MoveJ (P_Roof_J_p02_w05)
  MoveJ (P_Roof_J_p02_w06)
  MoveJ (P_Roof_J_p03_w00)
  MoveJ (P_Roof_J_p03_w01)
  MoveJ (P_Roof_J_p03_w02)
  MoveJ (P_Roof_J_p03_w03)
  MoveJ (P_Roof_J_p03_w04)
  MoveJ (P_Roof_J_p03_w05)
  MoveJ (P_Roof_J_p03_w06)
  MoveJ (P_Roof_J_p04_w00)
  MoveJ (P_Roof_J_p04_w01)
  MoveJ (P_Roof_J_p04_w02)
  MoveJ (P_Roof_J_p04_w03)
  MoveJ (P_Roof_J_p04_w04)
  MoveJ (P_Roof_J_p04_w05)
  MoveJ (P_Roof_J_p04_w06)
  MoveJ (P_Roof_J_p05_w00)
  MoveJ (P_Roof_J_p05_w01)
  MoveJ (P_Roof_J_p05_w02)
  MoveJ (P_Roof_J_p05_w03)
  MoveJ (P_Roof_J_p05_w04)
  MoveJ (P_Roof_J_p05_w05)
  MoveJ (P_Roof_J_p05_w06)
  MoveJ (P_Home)

--- program Paint_Hood (robot Comau Smart5 NJ 130-2.6) ---
  Set Ref.: CarFrame
  Set Tool: Generic Paint Sprayer
  MoveJ (P_Home)
  MoveJ (P_Hood_J_approach)
  MoveJ (P_Hood_J_p00_w00)
  MoveJ (P_Hood_J_p00_w01)
  MoveJ (P_Hood_J_p00_w02)
  MoveJ (P_Hood_J_p00_w03)
  MoveJ (P_Hood_J_p00_w04)
  MoveJ (P_Hood_J_p01_w00)
  MoveJ (P_Hood_J_p01_w01)
  MoveJ (P_Hood_J_p01_w02)
  MoveJ (P_Hood_J_p01_w03)
  MoveJ (P_Hood_J_p01_w04)
  MoveJ (P_Hood_J_p02_w00)
  MoveJ (P_Hood_J_p02_w01)
  MoveJ (P_Hood_J_p02_w02)
  MoveJ (P_Hood_J_p02_w03)
  MoveJ (P_Hood_J_p02_w04)
  MoveJ (P_Hood_J_p03_w00)
  MoveJ (P_Hood_J_p03_w01)
  MoveJ (P_Hood_J_p03_w02)
  MoveJ (P_Hood_J_p03_w03)
  MoveJ (P_Hood_J_p03_w04)
  MoveJ (P_Hood_J_p04_w00)
  MoveJ (P_Hood_J_p04_w01)
  MoveJ (P_Hood_J_p04_w02)
  MoveJ (P_Hood_J_p04_w03)
  MoveJ (P_Hood_J_p04_w04)
  MoveJ (P_Home)

--- program Paint_Trunk (robot Comau Smart5 NJ 130-2.6) ---
  Set Ref.: CarFrame
  Set Tool: Generic Paint Sprayer
  MoveJ (P_Home)
  MoveJ (P_Trunk_J_approach)
  MoveJ (P_Trunk_J_p00_w00)
  MoveJ (P_Trunk_J_p00_w01)
  MoveJ (P_Trunk_J_p00_w02)
  MoveJ (P_Trunk_J_p00_w03)
  MoveJ (P_Trunk_J_p00_w04)
  MoveJ (P_Trunk_J_p01_w00)
  MoveJ (P_Trunk_J_p01_w01)
  MoveJ (P_Trunk_J_p01_w02)
  MoveJ (P_Trunk_J_p01_w03)
  MoveJ (P_Trunk_J_p01_w04)
  MoveJ (P_Trunk_J_p02_w00)
  MoveJ (P_Trunk_J_p02_w01)
  MoveJ (P_Trunk_J_p02_w02)
  MoveJ (P_Trunk_J_p02_w03)
  MoveJ (P_Trunk_J_p02_w04)
  MoveJ (P_Trunk_J_p03_w00)
  MoveJ (P_Trunk_J_p03_w01)
  MoveJ (P_Trunk_J_p03_w02)
  MoveJ (P_Trunk_J_p03_w03)
  MoveJ (P_Trunk_J_p03_w04)
  MoveJ (P_Trunk_J_p04_w00)
  MoveJ (P_Trunk_J_p04_w01)
  MoveJ (P_Trunk_J_p04_w02)
  MoveJ (P_Trunk_J_p04_w03)
  MoveJ (P_Trunk_J_p04_w04)
  MoveJ (P_Trunk_J_p05_w00)
  MoveJ (P_Trunk_J_p05_w01)
  MoveJ (P_Trunk_J_p05_w02)
  MoveJ (P_Trunk_J_p05_w03)
  MoveJ (P_Trunk_J_p05_w04)
  MoveJ (P_Trunk_J_p06_w00)
  MoveJ (P_Trunk_J_p06_w01)
  MoveJ (P_Trunk_J_p06_w02)
  MoveJ (P_Trunk_J_p06_w03)
  MoveJ (P_Trunk_J_p06_w04)
  MoveJ (P_Trunk_J_p07_w00)
  MoveJ (P_Trunk_J_p07_w01)
  MoveJ (P_Trunk_J_p07_w02)
  MoveJ (P_Trunk_J_p07_w03)
  MoveJ (P_Trunk_J_p07_w04)
  MoveJ (P_Home)
